(* IEC 61131-3 sources: Gen-AI/docs/member2_validation/codesys_release_v1.1/task_S07_skeleton, 1 file *)

(* ---- source.st ---- *)
FUNCTION_BLOCK FB_S07
VAR_INPUT
    BottleIn : BOOL;
    FillDone : BOOL;
    CapDone : BOOL;
    PackDone : BOOL;
    StartBtn : BOOL;
    EStop_NC : BOOL;
END_VAR
VAR_OUTPUT
    Conveyor : BOOL;
    FillValve : BOOL;
    CapMotor : BOOL;
    PackCyl : BOOL;
    CycleCount : UINT;
    Status : WORD;
END_VAR
(* Add a VAR block for internal state/timers before the implementation, if needed. *)
(* SKELETON ONLY: replace this RETURN with scan logic and required initial state. *)
RETURN;
END_FUNCTION_BLOCK
